Staubli VAL3: selEndProg.pgx

public program selEndProg()
begin
  nProgType=1
end
